Fanuc KAREL source: IO0196.KL

PROGRAM IO0196
%NOLOCKGROUP
%ENVIRONMENT REGOPE
ROUTINE RTEST
VAR
  I : INTEGER
  STATUS : INTEGER
  ENTRY : INTEGER
  A : ARRAY[3] OF INTEGER
  B : BOOLEAN
  R : REAL
  P : XYZWPR
  JPOS : JOINTPOS
  PF : POSITION
BEGIN
  I = 1
  A[1] = 2
  B = TRUE
  R = 1.0
  P = GET_POS_REG(1,STATUS,1)
  IF P.X > 0.0 THEN
    I = I + 1
  ENDIF
END RTEST
BEGIN
  RTEST
END IO0196
